(* IEC 61131-3 sources: beckhoffAutomationInterface/ST/VariantSample, 4 files *)

(* ---- GVL_MachineConfig.st ---- *)
(* The only file that names machines. Every other POU reads these constants
   or tests a feature define (PCV_MODBUS / PCV_ETHERCAT), never a machine name. *)
{attribute 'qualified_only'}
VAR_GLOBAL CONSTANT
{IF defined (MachineA)}
    MACHINE_NAME     : STRING(16) := 'MachineA';
    MAX_PRESSURE_BAR : REAL       := 3.0;
    DOORS_FITTED     : BOOL       := FALSE;
{ELSIF defined (MachineB)}
    MACHINE_NAME     : STRING(16) := 'MachineB';
    MAX_PRESSURE_BAR : REAL       := 10.0;
    DOORS_FITTED     : BOOL       := TRUE;
{END_IF}
END_VAR

(* ---- MAIN.st ---- *)
PROGRAM MAIN
VAR
    sMachine     : STRING(16);
    rMaxPressure : REAL;
    bDoorsFitted : BOOL;
    sPcvDriver   : STRING(16);
END_VAR

{IF defined (MachineA)}
{warning 'VARIANT CHECK: MachineA branch compiled'}
{ELSIF defined (MachineB)}
{warning 'VARIANT CHECK: MachineB branch compiled'}
{ELSE}
{error 'No machine variant selected (MachineA or MachineB)'}
{END_IF}

// Values: plain constants from the machine configuration.
sMachine     := GVL_MachineConfig.MACHINE_NAME;
rMaxPressure := GVL_MachineConfig.MAX_PRESSURE_BAR;
bDoorsFitted := GVL_MachineConfig.DOORS_FITTED;

// Structure: a feature define selects the driver.
{IF defined (PCV_MODBUS)}
{warning 'FEATURE CHECK: PCV_MODBUS driver compiled'}
PRG_PcvModbus();
sPcvDriver := PRG_PcvModbus.sName;
{ELSIF defined (PCV_ETHERCAT)}
{warning 'FEATURE CHECK: PCV_ETHERCAT driver compiled'}
PRG_PcvEtherCAT();
sPcvDriver := PRG_PcvEtherCAT.sName;
{ELSE}
{error 'No PCV feature selected (PCV_MODBUS or PCV_ETHERCAT)'}
{END_IF}

(* ---- PRG_PcvEtherCAT.st ---- *)
PROGRAM PRG_PcvEtherCAT
VAR_OUTPUT
    sName : STRING(16) := 'EtherCAT';
END_VAR
VAR
    nCycles : UDINT;
END_VAR

nCycles := nCycles + 1;

(* ---- PRG_PcvModbus.st ---- *)
PROGRAM PRG_PcvModbus
VAR_OUTPUT
    sName : STRING(16) := 'Modbus';
END_VAR
VAR
    nCycles : UDINT;
END_VAR

nCycles := nCycles + 1;
